// TIA Portal V20 export
// export: Created 2026-10-12T16:46:22.7082025Z, ExportSetting WithDefaults, DisplayName Totally Integrated Automation Portal, DisplayVersion V20 Update 6, DisplayName TIA Portal Openness, DisplayVersion V20 Update 6, DisplayName TIA Portal Version Control Interface, DisplayVersion V20 Update 6, DisplayName SINAMICS Startdrive Advanced, DisplayVersion V20 SP1 Update 2, DisplayName SINAMICS Startdrive G110M, G120, G120C, G120D, G120P, G115D, DisplayVersion V20 SP1 Update 2, DisplayName SINAMICS Startdrive G130, G150, S120, S150, SINAMICS MV, G220, S200, S210, DisplayVersion V20 SP1 Update 2, DisplayName STEP 7 Professional, DisplayVersion V20 Update 6, DisplayName STEP 7 Safety, DisplayVersion V20 Update 2, DisplayName WinCC Basic/Comfort/Advanced, DisplayVersion V20 Update 6, DisplayName WinCC Professional, DisplayVersion V20 Update 6, DisplayName WinCC Unified, DisplayVersion V20 Update 6
TYPE "UDT_FK_OUT"
// stored: IsFailsafeCompliant false
   STRUCT
      PageNo : Word;   // Byte 0-1: imer 0
      Control : Word;   // Byte 2-3: 0=Aus, 3=Ein+Start
      SetVoltage : Int;   // Byte 4-5: x0.01V
      setCurrent : Int;   // Byte 6-7: x1A
      Reserved : Array[0..7] of Word;   // Byte 8-23: ungenutzt
      Padding : Array[0..3] of Word;   // Byte 24-31: ungenutzt
   END_STRUCT;
END_TYPE
